Fanuc KAREL source: kt00080.KL

-- PROVISIONAL review KL for V770-1; original PC SHA256 42befe0b5df7633f16ee15ec339d41655a322c2eea0d1e4d6bc205c66f7a1512
-- Incomplete behavior may be omitted. Consult companion uncertainty JSON. Do not deploy.
PROGRAM KT00080
%NOLOCKGROUP
VAR
  R1 : REAL
  OUT : REAL
-- UNRESOLVED_DECL H2 type=002017
BEGIN
  -- UNRESOLVED_PC offsets 5-16; opcodes 2E,23
  -- UNRESOLVED_PC offsets 21-35; opcodes 2E,22,9D,33,B4
  -- UNRESOLVED_PC offsets 40-63; opcodes 21,22,9D,33,B3,64,6B,23
  -- UNRESOLVED_PC offsets 68-72; opcodes 7F
END KT00080
